(* IEC 61131-3 sources: llm-plc-st-eval/data/processed_definitivo/gemini-3.1-pro-preview/A3/zero_shot, 3 files *)

(* ---- ejec_1.st ---- *)
FUNCTION_BLOCK FB_Com
VAR_INPUT
    txReq : BOOL;   // Petición de transmisión
    rxOk : BOOL;    // Confirmación de recepción
    rxData : INT;   // Dato recibido
END_VAR

VAR_OUTPUT
    txData : INT;   // Dato a transmitir
    ocupado : BOOL; // Intercambio en curso
    ok : BOOL;      // Intercambio exitoso
    error : BOOL;   // Intercambio fallido tras 3 intentos
    nIntentos : INT;// Número de intento actual (1, 2 o 3)
END_VAR

VAR
    rtTxReq : R_TRIG; // Detector de flanco para txReq
    rtRxOk : R_TRIG;  // Detector de flanco para rxOk
    timer : TON;      // Temporizador de 500ms
    timerIn : BOOL;   // Control de inicio/reinicio del temporizador
END_VAR

// Detección de flancos ascendentes
rtTxReq(CLK := txReq);
rtRxOk(CLK := rxOk);

// Inicio de un nuevo intercambio (se ignora si ya está ocupado)
IF rtTxReq.Q AND NOT ocupado THEN
    txData := 100;
    ocupado := TRUE;
    ok := FALSE;
    error := FALSE;
    nIntentos := 1;
    timerIn := FALSE; // Fuerza un ciclo en FALSE para reiniciar el temporizador
END_IF;

// Actualización del temporizador
timer(IN := timerIn, PT := T#500MS);

// Máquina de estados durante el intercambio
IF ocupado THEN
    IF timerIn THEN
        // El temporizador está corriendo, evaluar condiciones de respuesta o timeout
        IF rtRxOk.Q AND (rxData = txData) THEN
            // Éxito: se recibió confirmación con el eco correcto
            ok := TRUE;
            ocupado := FALSE;
            timerIn := FALSE;

        ELSIF timer.Q OR (rtRxOk.Q AND (rxData <> txData)) THEN
            // Falla: por tiempo agotado o por dato incorrecto
            IF nIntentos < 3 THEN
                nIntentos := nIntentos + 1;
                timerIn := FALSE; // Reinicia el temporizador en el próximo ciclo
            ELSE
                // Fallaron los 3 intentos permitidos
                error := TRUE;
                ocupado := FALSE;
                timerIn := FALSE;
            END_IF;
        END_IF;
    ELSE
        // Activar el temporizador para iniciar el conteo del intento actual
        timerIn := TRUE;
    END_IF;
ELSE
    // Asegurar que el temporizador se mantenga apagado si no hay intercambio activo
    timerIn := FALSE;
END_IF;
END_FUNCTION_BLOCK

(* ---- ejec_2.st ---- *)
FUNCTION_BLOCK FB_Com
VAR_INPUT
    txReq : BOOL;
    rxOk : BOOL;
    rxData : INT;
END_VAR
VAR_OUTPUT
    txData : INT;
    ocupado : BOOL;
    ok : BOOL;
    error : BOOL;
    nIntentos : INT;
END_VAR
VAR
    txReq_Trig : R_TRIG;
    rxOk_Trig : R_TRIG;
    temporizador : TON;
    estado : INT := 0; // 0: Reposo, 1: Intercambio en curso
END_VAR

// Detección de flancos ascendentes
txReq_Trig(CLK := txReq);
rxOk_Trig(CLK := rxOk);

// Actualización del temporizador
temporizador(IN := (estado = 1), PT := T#500MS);

CASE estado OF
    0: // Reposo: esperando nueva petición
        IF txReq_Trig.Q THEN
            txData := 100;
            ocupado := TRUE;
            ok := FALSE;
            error := FALSE;
            nIntentos := 1;
            estado := 1;

            // Reinicio forzado del temporizador para el intento 1
            temporizador(IN := FALSE);
            temporizador(IN := TRUE, PT := T#500MS);
        END_IF;

    1: // Intercambio en curso: esperando respuesta o timeout
        IF rxOk_Trig.Q THEN
            IF rxData = txData THEN
                // Éxito: confirmación recibida con eco correcto
                ok := TRUE;
                ocupado := FALSE;
                estado := 0;
            ELSE
                // Fallo: confirmación recibida pero dato incorrecto
                nIntentos := nIntentos + 1;
                temporizador(IN := FALSE);
                temporizador(IN := TRUE, PT := T#500MS);
            END_IF;
        ELSIF temporizador.Q THEN
            // Fallo: vencimiento del plazo de 500 ms sin confirmación
            nIntentos := nIntentos + 1;
            temporizador(IN := FALSE);
            temporizador(IN := TRUE, PT := T#500MS);
        END_IF;

        // Evaluación del límite máximo de intentos
        IF estado = 1 AND nIntentos > 3 THEN
            error := TRUE;
            ocupado := FALSE;
            nIntentos := 3; // Conserva el último valor válido
            estado := 0;
        END_IF;
END_CASE;
END_FUNCTION_BLOCK

(* ---- ejec_3.st ---- *)
FUNCTION_BLOCK FB_Com
VAR_INPUT
    txReq : BOOL;
    rxOk : BOOL;
    rxData : INT;
END_VAR
VAR_OUTPUT
    txData : INT;
    ocupado : BOOL;
    ok : BOOL;
    error : BOOL;
    nIntentos : INT;
END_VAR
VAR
    reqTrig : R_TRIG;
    rxTrig : R_TRIG;
    timer : TON;
END_VAR

// Detectar flancos de subida en las señales de control
reqTrig(CLK := txReq);
rxTrig(CLK := rxOk);

// Iniciar un nuevo intercambio (se ignora si ya está en curso)
IF reqTrig.Q AND NOT ocupado THEN
    txData := 100;
    ocupado := TRUE;
    ok := FALSE;
    error := FALSE;
    nIntentos := 1;
    timer(IN := FALSE, PT := T#500MS); // Reset inicial del temporizador
END_IF;

// Lógica de control durante el intercambio activo
IF ocupado THEN
    // Ejecutar temporizador para el intento actual
    timer(IN := TRUE, PT := T#500MS);

    // Evaluar si se recibe confirmación con el dato correcto (eco)
    IF rxTrig.Q AND (rxData = txData) THEN
        ok := TRUE;
        ocupado := FALSE;
        timer(IN := FALSE, PT := T#500MS); // Detener temporizador

    // Evaluar si el intento falla (por timeout o por dato incorrecto)
    ELSIF timer.Q OR (rxTrig.Q AND (rxData <> txData)) THEN
        IF nIntentos < 3 THEN
            nIntentos := nIntentos + 1;        // Incrementar contador de intentos
            timer(IN := FALSE, PT := T#500MS); // Reiniciar temporizador para el nuevo intento
        ELSE
            error := TRUE;                     // Activar error tras agotar los 3 intentos
            ocupado := FALSE;
            timer(IN := FALSE, PT := T#500MS); // Detener temporizador
        END_IF;
    END_IF;
ELSE
    // Mantener el temporizador inactivo cuando no hay intercambio
    timer(IN := FALSE, PT := T#500MS);
END_IF;
END_FUNCTION_BLOCK
